// TIA Portal V21 export
// export: Created 2026-11-11T00:47:39.6596702Z, ExportSetting WithDefaults, DisplayName Totally Integrated Automation Portal, DisplayVersion V21 Update 3, DisplayName STEP 7 Professional, DisplayVersion V21 Update 3, DisplayName STEP 7 Safety, DisplayVersion V21, DisplayName Tech WebApplication, DisplayVersion V21, DisplayName WinCC Basic/Comfort/Advanced, DisplayVersion V21 Update 3, DisplayName WinCC Unified, DisplayVersion V21 Update 3
FUNCTION_BLOCK "FB_Fbd_ex150"   // FB158, FBD
{ S7_Optimized_Access := 'TRUE' }
VERSION : 0.1
// stored: AutoNumber true, IsIECCheckEnabled false, IsRetainMemResEnabled false, MemoryReserve 100, SetENOAutomatically false, UDAEnableTagReadback false
   VAR_INPUT
      v_req : Bool;
      v_db_number : DB_ANY;
   END_VAR
   VAR_OUTPUT
      v_ret_val : Int;
      v_db_length : UDInt;
      v_attrib : Byte;
   END_VAR
BEGIN

REGION Network 1: ATTR_DB - Read data block attribute
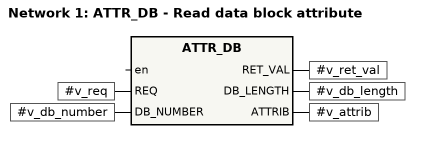
   #v_ret_val := ATTR_DB(REQ := #v_req,
                         DB_NUMBER := #v_db_number,
                         DB_LENGTH => #v_db_length,
                         ATTRIB => #v_attrib);
END_REGION
END_FUNCTION_BLOCK
